KUKA KRL program: WeldPair1.src

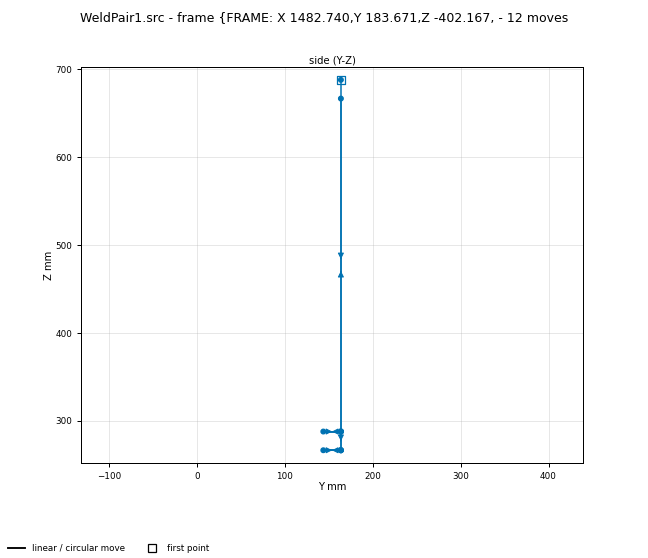
[picture p0: tool path of WeldPair1.src in frame {FRAME: X 1482.740,Y 183.671,Z -402.167,, 12 of 13 moves have a stored position in this frame; points joined in program order, loops and branches not executed]
&ACCESS RVP
&REL 1
&PARAM TEMPLATE = C:\KRC\Roboter\Template\vorgabe
&PARAM EDITMASK = *
DEF WeldPair1 ( )

; External program calls:
EXT DoWeld()

EXT BAS (BAS_COMMAND :IN,REAL :IN )


; GLOBAL INTERRUPT DECL 3 WHEN $STOPMESS==TRUE DO IR_STOPM ( )
; INTERRUPT ON 3

;FOLD Initialise and set default speed
BAS (#INITMOV,0)
BAS (#VEL_PTP,100)
BAS (#ACC_PTP,20)
$VEL.CP=0.2
BAS (#TOOL,0)
BAS (#BASE,0)
;ENDFOLD

;;FOLD STARTPOS
;$BWDSTART = FALSE
;PDAT_ACT = PDEFAULT
;BAS(#PTP_DAT)
;FDAT_ACT = {TOOL_NO 0,BASE_NO 0,IPO_FRAME #BASE}
;BAS(#FRAMES)
;;ENDFOLD

$ADVANCE = 5

;FOLD ---- Quickly skip BCO ----
; PTP $AXIS_ACT
;ENDFOLD

;FOLD ---- GO HOME ----
; PTP {A1 0.000, A2 -90.000, A3 90.000, A4 0.000, A5 0.000, A6 0.000, E1 0, E2 0, E3 0, E4 0, E5 0, E6 0}
;ENDFOLD


; Program generated by VerticalBot Studio for KUKA KR 120 R2900 extra on 25/10/2026 12:00:00
; Using nominal kinematics.
; ---- Setting reference (Base) ----
$BASE = {FRAME: X 1482.740,Y 183.671,Z -402.167,A 6.534,B 0.000,C 0.000}
; --------------------------
; ---- Setting tool (TCP) ----
$TOOL = {FRAME: X 0.270,Y 0.000,Z 1049.990,A 0.000,B -90.000,C 0.000}
; --------------------------
; show WeldGun
$VEL.CP = 1.00000
PTP {A1 -12.43810,A2 -78.90300,A3 98.90130,A4 -0.00000,A5 70.00160,A6 -95.90410}
LIN {X 220.309,Y 163.798,Z 688.010,A -90.000,B 90.000,C 0.000}
LIN {X 220.309,Y 163.798,Z 288.010,A -90.000,B 90.000,C 0.000}
LIN {X 220.309,Y 163.798,Z 288.010,A -90.000,B 90.000,C 0.000}
LIN {X 220.309,Y 163.798,Z 288.010,A -90.000,B 90.000,C 0.000}
$VEL.CP = 0.05000
LIN {X 220.309,Y 143.798,Z 288.010,A -90.000,B 90.000,C 0.000}
DoWeld(10)
LIN {X 220.309,Y 163.798,Z 288.010,A -90.000,B 90.000,C 0.000}
$VEL.CP = 1.00000
LIN {X 220.309,Y 163.798,Z 266.723,A -90.000,B 90.000,C 0.000}
$VEL.CP = 0.05000
LIN {X 220.309,Y 143.798,Z 266.723,A -90.000,B 90.000,C 0.000}
DoWeld()
LIN {X 220.309,Y 163.798,Z 266.723,A -90.000,B 90.000,C 0.000}
$VEL.CP = 1.00000
LIN {X 220.309,Y 163.798,Z 266.723,A -90.000,B 90.000,C 0.000}
LIN {X 220.309,Y 163.798,Z 266.723,A -90.000,B 90.000,C 0.000}
LIN {X 220.309,Y 163.798,Z 666.723,A -90.000,B 90.000,C 0.000}
END
